# EPICS substitutions: db/Beckhoff_7XXX/ecmcEP7211-0034_OPT_cst.substitutions
file "ecmcEL72XX_DRV_CST.template"
{
  pattern {CH_ID, ESLO, EGU}
          {01,    0.1,  "%"}
}

file "ecmc_analogInput-chX.template"
{
  pattern {CH_ID, sourceName,       KEY,   suffix,    DESC,         EGU,     ESLO,      PREC, LOPR, HOPR, LOLO, LOW, HIGH, HIHI, HYST, LLSV,       LSV,        HSV,        HHSV}
          {01,    "velocityActual", "Drv", "-VelAct", "Actual Vel", "rad/s", 2.3406E-5, 3,    0,    0,    0,    0,   0,    0,    0,    "NO_ALARM", "NO_ALARM", "NO_ALARM", "NO_ALARM"}
          {01,    "infoData",       "Drv", "-VolAct", "InfoData1",  "V",     0.001,     1,    0,    60,   8,    20,  49,   50,   0.25, "MAJOR",    "MINOR",    "MINOR",    "MAJOR"}
}

file "ecmcEL72XX_FB_STAT.template"
{
  pattern {CH_ID}
          {01   }
}
